Fanuc KAREL source: KT00773.KL

PROGRAM KT00773
%NOLOCKGROUP
VAR
  I1: INTEGER
  I2: INTEGER
  OUT: REAL
BEGIN
  I1 = 2
  I2 = 3
  I1 = 2
  I2 = 3
  OUT = ASIN(I1)
END KT00773
